{attribute 'qualified_only' := ''}
{attribute 'strict' := ''}
TYPE E_SplineType :
(
	SPLINE_NATURAL := 0,
	SPLINE_FIXEDBOUNDARY := 1,
	SPLINE_NONODEBOUNDARY := 2
);
END_TYPE

(* stored: Version 1.1.0.1, ProductVersion 3.1.4024.12
   DUT E_SplineType: Id {7989b57e-1a9f-405d-9359-f5e4387b39ee} *)
